(* IEC 61131-3 sources: garage-sweeper/PLC/src/Contracts, 8 files *)

(* ---- HmiCommand.st ---- *)
TYPE HmiCommand :
STRUCT
	sequence : UDINT;
	code : HmiCommandCode;
	manualTwist : Twist;
END_STRUCT
END_TYPE

(* ---- HmiCommandCode.st ---- *)
{attribute 'qualified_only'}
{attribute 'strict'}
TYPE HmiCommandCode :
(
	NONE := 0,
	MANUAL_DRIVE,
	START_MAPPING,
	START_SWEEPING,
	PAUSE,
	RESUME,
	STOP,
	GO_TO_DOCK,
	EMERGENCY_STOP,
	RESET
) INT;
END_TYPE

(* ---- HmiStatus.st ---- *)
TYPE HmiStatus :
STRUCT
	acknowledgedSequence : UDINT;
	missionState : MissionState;
	lastRejection : STRING(80);
	estimatedPose : Pose2D;
	isSimulatorConnected : BOOL;
	isLidarOk : BOOL;
	hasMap : BOOL;
END_STRUCT
END_TYPE

(* ---- MissionState.st ---- *)
{attribute 'qualified_only'}
{attribute 'strict'}
TYPE MissionState :
(
	IDLE := 0,
	MANUAL,
	MAPPING,
	SWEEPING,
	PAUSED,
	RETURNING_TO_DOCK,
	DOCKED,
	EMERGENCY_STOPPED
) INT;
END_TYPE

(* ---- SimulatorCommand.st ---- *)
TYPE SimulatorCommand :
STRUCT
	version : UDINT;
	cycle : UDINT;
	plcTimeInNs : ULINT;
	// The wheels' actual speed, from the NC axes. The simulator moves the robot with it.
	leftWheelVelocityInMPerS : LREAL;
	rightWheelVelocityInMPerS : LREAL;
	isLeftDriveEnabled : BOOL;
	isRightDriveEnabled : BOOL;
	isLidarPowered : BOOL;
	estimatedPose : Pose2D;
END_STRUCT
END_TYPE

(* ---- SimulatorFeedback.st ---- *)
TYPE SimulatorFeedback :
STRUCT
	version : UDINT;
	sequence : UDINT;
	timeInNs : ULINT;
	leftWheelAngleInRad : LREAL;
	rightWheelAngleInRad : LREAL;
	leftWheelVelocityInRadPerS : LREAL;
	rightWheelVelocityInRadPerS : LREAL;
	angularRateInRadPerS : Vector3;
	accelerationInMPerS2 : Vector3;
	truePose : Pose2D;
	collided : BOOL;
END_STRUCT
END_TYPE

(* ---- RobotHmi.st ---- *)
{attribute 'qualified_only'}
VAR_GLOBAL
	command : HmiCommand;
	status : HmiStatus;
END_VAR

(* ---- SimulatorIo.st ---- *)
{attribute 'qualified_only'}
VAR_GLOBAL
	command : SimulatorCommand;
	feedback : SimulatorFeedback;
	scan : LaserScan;
END_VAR
